(* IEC 61131-3 sources: plc-iiot-stack/flagship/src/POUs/Iiot/PRG_Iiot, 5 files *)

(* ---- FillNodePoints.method.impl.st ---- *)
IF ltNow >= ltStart THEN
    aPoints[GVL_IiotMap.PT_PLC1_UPTIME].lrValue := ULINT_TO_LREAL(LTIME_TO_ULINT(ltNow - ltStart) / NS_PER_S);
END_IF
IF fbDiag.udiConnects > 0 THEN
    aPoints[GVL_IiotMap.PT_PLC1_RECONNECTS].lrValue := UDINT_TO_LREAL(fbDiag.udiConnects - 1);
END_IF
aPoints[GVL_IiotMap.PT_PLC1_QUEUE].lrValue := UINT_TO_LREAL(fbTelemetry.uiPending + fbAlarms.uiPending);
aPoints[GVL_IiotMap.PT_PLC1_DROPPED].lrValue :=
    UDINT_TO_LREAL(fbTelemetry.udiDropped + fbAlarms.udiDropped + fbCommands.udiAckFailed);
aPoints[GVL_IiotMap.PT_PLC1_CMD_ACCEPTED].lrValue := UDINT_TO_LREAL(fbCommands.udiAccepted);
aPoints[GVL_IiotMap.PT_PLC1_CMD_REJECTED].lrValue := UDINT_TO_LREAL(fbCommands.udiRejected + fbCommands.udiDropped);
aPoints[GVL_IiotMap.PT_PLC1_UPTIME].eQuality := E_IiotQuality.Good;
aPoints[GVL_IiotMap.PT_PLC1_RECONNECTS].eQuality := E_IiotQuality.Good;
aPoints[GVL_IiotMap.PT_PLC1_QUEUE].eQuality := E_IiotQuality.Good;
aPoints[GVL_IiotMap.PT_PLC1_DROPPED].eQuality := E_IiotQuality.Good;
aPoints[GVL_IiotMap.PT_PLC1_CMD_ACCEPTED].eQuality := E_IiotQuality.Good;
aPoints[GVL_IiotMap.PT_PLC1_CMD_REJECTED].eQuality := E_IiotQuality.Good;

(* ---- PRG_Iiot.decl.st ---- *)
// Назначение: ПЛК-часть IIoT-стека во флагмане КНС-1: связь с брокером и состояние узла (FB_MqttDiag),
//             телеметрия (FB_MqttTelemetry), тревоги (FB_MqttAlarms) и шлюз команд (FB_MqttCommands) поверх
//             переменных флагмана: значения и слова тревог устройств и станции читает, а принятые команды
//             пишет FB_IiotKnsMap (сгенерирован из schema/). Таблицы метрик, команд и тревог — GVL_IiotMap.
//             Клиент MQTT — itfClientOverride (адаптер библиотеки) или FB_MqttClientNone. Задача MainTask
//             флагмана, после PRG_Devices. Настройки — GVL_Iiot.stIiotCfg, состояние — GVL_Iiot.stIiotSts.
// Автор:      kr0nsch
// Версия:     0.2.0
// Документ:   docs/plc_mqtt.md, раздел «Привязка к флагману»
PROGRAM PRG_Iiot
VAR_INPUT
    itfClientOverride : I_MqttClient;     // адаптер библиотеки или подменный клиент; 0 — FB_MqttClientNone
END_VAR
VAR
    fbClientNone : FB_MqttClientNone;
    itfClient : I_MqttClient;
    fbMap : FB_IiotKnsMap;
    fbDiag : FB_MqttDiag;
    fbTelemetry : FB_MqttTelemetry;
    fbAlarms : FB_MqttAlarms;
    fbCommands : FB_MqttCommands;
    aPoints : ARRAY[1..GVL_IiotMap.POINT_COUNT] OF ST_IiotPoint;
    aAlarms : ARRAY[1..GVL_IiotMap.ALARM_COUNT] OF ST_IiotAlarm;
    aAlarmWords : ARRAY[1..GVL_IiotMap.ALARM_WORDS_COUNT] OF ST_IiotAlarmWords;
    aRules : ARRAY[1..GVL_IiotMap.RULE_COUNT] OF ST_IiotCmdRule;
    xInitDone : BOOL;
    ltStart : LTIME;                      // первый вызов: отсчёт uptime
    ltNow : LTIME;
    uliTs_ms : ULINT;
    xClockValid : BOOL;
    sPrefix : STRING(GVL_Const.IIOT_PREFIX_LEN);
    uiDevSeq : UINT;
    iDevResult : INT;
    diIdx : DINT;
END_VAR
VAR CONSTANT
    RTC_OK : UDINT := 0;                  // SysTimeRtcHighResGet: «нет ошибки» (ERR_OK)
    NS_PER_S : ULINT := 1000000000;
END_VAR

(* ---- PRG_Iiot.impl.st ---- *)
// 0. Таблицы настроек из схемы данных — один раз
ltNow := F_IiotNow();
IF NOT xInitDone THEN
    FOR diIdx := 1 TO GVL_IiotMap.POINT_COUNT DO
        aPoints[diIdx].stCfg := GVL_IiotMap.POINT_CFG[diIdx];
    END_FOR
    FOR diIdx := 1 TO GVL_IiotMap.ALARM_COUNT DO
        aAlarms[diIdx].stCfg := GVL_IiotMap.ALARM_CFG[diIdx];
    END_FOR
    FOR diIdx := 1 TO GVL_IiotMap.RULE_COUNT DO
        aRules[diIdx] := GVL_IiotMap.RULE_CFG[diIdx];
    END_FOR
    ltStart := ltNow;
    xInitDone := TRUE;
END_IF

// 1. Клиент MQTT: адаптер библиотеки (или подменный клиент тестов) либо клиент без транспорта
IF itfClientOverride <> 0 THEN
    itfClient := itfClientOverride;
ELSE
    itfClient := fbClientNone;
END_IF
itfClient.Cycle();

// 2. Время: монотонное — для таймаутов и периодов, календарное (UTC, мс) — для ts и проверки команд
xClockValid := SysTimeRtcHighResGet(pTimestamp := uliTs_ms) = RTC_OK AND F_IiotClockValid(uliTs_ms := uliTs_ms);
sPrefix := CONCAT(CONCAT(GVL_Iiot.stIiotCfg.sSite, GVL_Const.TOPIC_SEPARATOR), GVL_Iiot.stIiotCfg.sArea);
sPrefix := CONCAT(CONCAT(sPrefix, GVL_Const.TOPIC_SEPARATOR), GVL_Iiot.stIiotCfg.sUnit);

// 3. Значения флагмана -> метрики и слова тревог; метрики узла
fbMap.FillPoints(aPointTable := aPoints);
fbMap.FillAlarmWords(aWordTable := aAlarmWords);
FillNodePoints();

// 4. Связь и состояние узла
fbDiag(xEnable := GVL_Iiot.stIiotCfg.xEnable,
       itfClient := itfClient,
       ltNow := ltNow,
       uliTs_ms := uliTs_ms,
       sTopicPrefix := sPrefix,
       sNode := GVL_Iiot.stIiotCfg.sNode,
       sSwVersion := GVL_Iiot.stIiotCfg.sSwVersion,
       tPeriod := GVL_Iiot.stIiotCfg.tTelemetryPeriod,
       udiPubFailed := fbTelemetry.udiFailed + fbAlarms.udiFailed,
       stBroker := GVL_Iiot.stIiotCfg.stBroker);

// 5. Телеметрия и тревоги — после рождения узла
fbTelemetry(xEnable := GVL_Iiot.stIiotCfg.xEnable,
            xReady := fbDiag.xReady,
            itfClient := itfClient,
            ltNow := ltNow,
            uliTs_ms := uliTs_ms,
            sTopicPrefix := sPrefix,
            tPeriod := GVL_Iiot.stIiotCfg.tTelemetryPeriod,
            aPoints := aPoints);
fbAlarms(xEnable := GVL_Iiot.stIiotCfg.xEnable,
         xReady := fbDiag.xReady,
         itfClient := itfClient,
         uliTs_ms := uliTs_ms,
         sTopicPrefix := sPrefix,
         aAlarms := aAlarms,
         aWords := aAlarmWords);

// 6. Команды: состояние устройства команды в обработке, приём, запись в GVL_Hmi
IF fbCommands.xPending THEN
    fbMap.DeviceCmdState(diDev := RuleDevice(diRule := fbCommands.stCmd.diRule), uiSeq => uiDevSeq,
                         iResult => iDevResult);
END_IF
fbCommands(xEnable := GVL_Iiot.stIiotCfg.xEnable AND GVL_Iiot.stIiotCfg.xCommandsEnable,
           itfClient := itfClient,
           ltNow := ltNow,
           uliTs_ms := uliTs_ms,
           sTopicPrefix := sPrefix,
           uiDevSeq := uiDevSeq,
           iDevResult := iDevResult,
           aRules := aRules);
IF fbCommands.xCmdValid THEN
    fbMap.DeviceCmdState(diDev := RuleDevice(diRule := fbCommands.stCmd.diRule), uiSeq => uiDevSeq,
                         iResult => iDevResult);
    fbMap.ApplyCommand(diRule := fbCommands.stCmd.diRule, rValue := fbCommands.stCmd.rValue);
    fbCommands.Arm(uiSeqBefore := uiDevSeq);
END_IF

// 7. Состояние для HMI и SCADA
GVL_Iiot.stIiotSts.eConnState := fbDiag.eState;
GVL_Iiot.stIiotSts.eNe107 := fbDiag.eNe107;
GVL_Iiot.stIiotSts.udiConnects := fbDiag.udiConnects;
GVL_Iiot.stIiotSts.udiDisconnects := fbDiag.udiDisconnects;
GVL_Iiot.stIiotSts.udiConnectFailures := fbDiag.udiConnectFailures;
GVL_Iiot.stIiotSts.diLastError := fbDiag.diLastError;
GVL_Iiot.stIiotSts.udiPublished := fbTelemetry.udiPublished + fbAlarms.udiPublished;
GVL_Iiot.stIiotSts.udiPublishFailed := fbTelemetry.udiFailed + fbAlarms.udiFailed;
GVL_Iiot.stIiotSts.uiQueue := fbTelemetry.uiPending + fbAlarms.uiPending;
GVL_Iiot.stIiotSts.udiDropped := fbTelemetry.udiDropped + fbAlarms.udiDropped + fbCommands.udiAckFailed;
GVL_Iiot.stIiotSts.udiCmdAccepted := fbCommands.udiAccepted;
GVL_Iiot.stIiotSts.udiCmdRejected := fbCommands.udiRejected + fbCommands.udiDropped;
GVL_Iiot.stIiotSts.eLastCmdReason := fbCommands.eLastReason;
GVL_Iiot.stIiotSts.xClockValid := xClockValid;

(* ---- RuleDevice.method.decl.st ---- *)
// Номер устройства строки белого списка (для FB_IiotKnsMap.DeviceCmdState); вне таблицы — 0.
METHOD PRIVATE RuleDevice : DINT
VAR_INPUT
    diRule : DINT;
END_VAR

(* ---- RuleDevice.method.impl.st ---- *)
IF diRule >= 1 AND diRule <= GVL_IiotMap.RULE_COUNT THEN
    RuleDevice := aRules[diRule].diDev;
END_IF
